Yaskawa INFORM job: SZLIF_SPAWU_TROJNIKA.JBI

/JOB
//NAME SZLIF_SPAWU_TROJNIKA
///FOLDERNAME TROJNIKI
//POS
///NPOS 0,0,0,4,0,0
///USER 10
///TOOL 17
///POSTYPE USER
///RECTAN
///RCONF 1,0,0,0,0,0,0,0,0,0,0,0,0,0,0,0,0,0,0,0,0,0,0,0
P00010=63.000,1.000,-2.000,-90.0000,-90.0000,90.0000
///USER 8
P00011=8.000,1.000,-2.000,-90.0000,-90.0000,90.0000
P00012=63.000,1.000,10.000,-90.0000,-90.0000,90.0000
///RCONF 0,0,0,0,0,0,0,0,0,0,0,0,0,0,0,0,0,0,0,0,0,0,0,0
P00013=8.000,1.000,10.000,-90.0000,-90.0000,90.0000
//INST
///DATE 2026/07/21 11:39
///ATTR SC,RW
///GROUP1 RB1
NOP
'FREZ TOOL 17: KROK SREDNICY
'I073 USTAWIA OPERATOR
'I070=120 DLA FREZA 12MM
SET I020 200
SET I120 1
CALL JOB:OBLICZ_SZLIF_TROJNIKA
'WEJSCIE NA PROMIEN 3MM
MOVL P010 V=I020 PL=0
*OBIEG
'JEDEN PELNY OBIEG
MOVC P010 V=I020 PL=1
MOVC P013 V=I020 PL=1
MOVC P012 V=I020 PL=1
MOVC P011 V=I020 PL=1
MOVC P010 V=I020 PL=0
'KONIEC PO OBIEGU DOCELOWYM
IFTHENEXP D074<D120
	 ADD I120 1
	 CALL JOB:OBLICZ_SZLIF_TROJNIKA
	'PROMIENIOWY DOJAZD DO OBIEGU
	 MOVL P010 V=I020 PL=0
	 JUMP *OBIEG
ENDIF
RET
END
